(* IEC 61131-3 sources: Lasal-MCP/examples/SampleSource/LASALScreenAdvancedSolution/LASALScreenAdvancedSolution/LASALScreenAdvacnedSolution/Stations/Terminal/HMI/Class/MyValues, 1 file *)

(* ---- MyValues.st ---- *)
(*!
<Class
	Name               = "MyValues"
	Revision           = "0.0"
	RealtimeTask       = "false"
	CyclicTask         = "false"
	BackgroundTask     = "false"
	Sigmatek           = "false"
	OSInterface        = "false"
	HighPriority       = "false"
	Automatic          = "false"
	UpdateMode         = "Prescan"
	SharedCommandTable = "true"
	Objectsize         = "(360,300)">
	<Channels>
		<Server Name="Active" Visualized="true" Initialize="true" DefValue="1" WriteProtected="false" Retentive="false"/>
		<Server Name="ID" Visualized="true" Initialize="true" WriteProtected="true" Retentive="false"/>
		<Server Name="Value1" Visualized="true" Initialize="true" DefValue="111" WriteProtected="false" Retentive="File"/>
		<Server Name="Value2" Visualized="true" Initialize="true" DefValue="222" WriteProtected="false" Retentive="File"/>
		<Server Name="Value3" Visualized="true" Initialize="true" DefValue="333" WriteProtected="false" Retentive="File"/>
	</Channels>
</Class>
*)
MyValues : CLASS
  //Servers:
	Value1 	: SvrChCmd_DINT;
	Value2 	: SvrCh_DINT;
	Value3 	: SvrCh_DINT;
	Active 	: SvrCh_DINT;
	ID 	: SvrCh_DINT;
  //Clients:
  //Variables:
  //Functions:
  //Tables:
	FUNCTION @STD
		VAR_OUTPUT
			ret_code	: CONFSTATES;
		END_VAR;
	FUNCTION GLOBAL TAB @CT_;
END_CLASS;
